TYPE "ST_UnitProbeStationCfg"
VERSION : 0.1
   STRUCT
      "SchemaVersion" : UInt := 1;
      "SiteLabel" : String[80] := 'bench';
      "Enabled" : Bool := TRUE;
   END_STRUCT;
END_TYPE
